// TIA Portal V21 export
TextList "TL_Cmd"  ListRange=Decimal
  TextListEntry   Text="-"
  TextListEntry   From=1, To=1, Text="1 PODIGNI"
  TextListEntry   From=2, To=2, Text="2 SPUSTI"
  TextListEntry   From=3, To=3, Text="3 POMAKNI"
  TextListEntry   From=10, To=10, Text="10 RESET"
